(* IEC 61131-3 sources: PLC-Static-Analysis/modules/plc-rules/src/test/resources/PLCA-Q001, 2 files *)

(* ---- compliant.st ---- *)
FUNCTION_BLOCK FB_Used
VAR
    nCount : INT;
    nForChildren : INT;
    aBuf : ARRAY[0..cMax] OF INT;
    nSpare1 : INT;
    bReserve_2 : BOOL;
    {attribute 'OPC.UA.DA' := '1'}
    rExposed : REAL;
    iSensor AT %I* : BOOL;
    pTarget : POINTER TO INT;
    nAddr : INT;
    nReadFromOutside : INT;
END_VAR
VAR CONSTANT
    cMax : INT := 9;
END_VAR
pTarget := ADR(nAddr);
aBuf[0] := 1;

METHOD Inc
nCount := nCount + 1;
END_METHOD
END_FUNCTION_BLOCK

FUNCTION_BLOCK FB_Child EXTENDS FB_Used
nForChildren := 0;
END_FUNCTION_BLOCK

FUNCTION_BLOCK ABSTRACT FB_Abstract_Base
VAR
    nForImplementations : INT;
END_VAR
END_FUNCTION_BLOCK

PROGRAM P_User
VAR
    fb : FB_Used;
    n : INT;
END_VAR
fb.Inc();
n := fb.nReadFromOutside;
END_PROGRAM

(* ---- noncompliant.st ---- *)
FUNCTION_BLOCK FB_Unused
VAR_INPUT
    bIn : BOOL;
END_VAR
VAR
    nNeverUsed : INT; // PLCA-Q001
    bUsed : BOOL;
    rTemp, rOther : REAL; // PLCA-Q001 PLCA-Q001
END_VAR
VAR_TEMP
    nScratch : DINT; // PLCA-Q001
END_VAR
bUsed := bIn;
END_FUNCTION_BLOCK

PROGRAM P_Main
VAR
    fbUnused : FB_Unused;
    fbNotCalled : FB_Unused; // PLCA-Q001
    n : INT;
END_VAR
fbUnused(bIn := n > 0);
END_PROGRAM

FUNCTION F_Unused : INT
VAR_INPUT
    nIn : INT;
END_VAR
VAR
    nLocal : INT; // PLCA-Q001
END_VAR
F_Unused := nIn;
END_FUNCTION
